{attribute 'qualified_only'}
{attribute 'strict'}
{attribute 'to_string'}
TYPE E_Tank_Target :
(
	eNone := 0,
	eClose,
	eOpen,
	eDrain,
	eClose_DrainPipe,
	eCIP
);
END_TYPE

(* stored: Version 1.1.0.1, ProductVersion 3.1.4024.12
   DUT E_Tank_Target: Id {15741c3f-3262-4749-a089-ec5958362e42} *)
